// TIA Portal V21 export
// export: Created 2026-11-11T00:47:16.600127Z, ExportSetting WithDefaults, DisplayName Totally Integrated Automation Portal, DisplayVersion V21 Update 3, DisplayName STEP 7 Professional, DisplayVersion V21 Update 3, DisplayName STEP 7 Safety, DisplayVersion V21, DisplayName Tech WebApplication, DisplayVersion V21, DisplayName WinCC Basic/Comfort/Advanced, DisplayVersion V21 Update 3, DisplayName WinCC Unified, DisplayVersion V21 Update 3
FUNCTION_BLOCK "FB_Fbd_ex043"   // FB86, FBD
{ S7_Optimized_Access := 'TRUE' }
VERSION : 0.1
// stored: AutoNumber true, IsIECCheckEnabled false, IsRetainMemResEnabled false, MemoryReserve 100, SetENOAutomatically false, UDAEnableTagReadback false
   VAR_INPUT
      v_part : PIP;
   END_VAR
   VAR_OUTPUT
      v_ret_val : Int;
      v_fladdr : Word;
   END_VAR
BEGIN

REGION Network 1: SYNC_PI - Synchronize the process image inputs
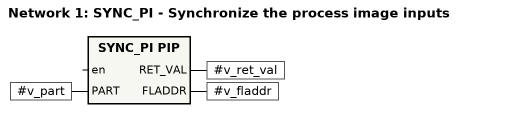
   #v_ret_val := SYNC_PI(PART := #v_part, FLADDR => #v_fladdr);
END_REGION
END_FUNCTION_BLOCK
